(*
SPDX-FileCopyrightText: © 2026 Oleksandr Tiutyk <trofimich@gmail.com>
SPDX-License-Identifier: MIT
License: https://opensource.org/license/mit
*)

(*!
<summary>Base class for one test whose body completes in a single PLC scheduling cycle.</summary>
<description>
Override ExecuteTest with the checks. Returning from the body completes the body automatically.
BeforeTest and AfterTest are optional scenario hooks. Constructor name identifies the case in reports.
Run through TestRunner, directly or inside a TestGroup. A complete run and its reporting may span more cycles
than the body. All instance access belongs to one task without reentry; other tasks need other instances.
</description>
*)

{attribute 'no_explicit_call' := 'do not call this function block directly'}
FUNCTION_BLOCK ABSTRACT SingleCycleTest EXTENDS TestCase

(*!
<summary>Implements the scenario body without runner guards or enumeration.</summary>
<description>
Keep persistent state in instance fields. Reporting a failure does not abort the current callback.
</description>
*)
METHOD PROTECTED ABSTRACT ExecuteTest
END_METHOD

(*!
<summary>Runs the body once and reports completion for the cycle.</summary>
*)
METHOD PROTECTED FINAL RunCycle : TEST_CYCLE_RESULT
ExecuteTest();
RunCycle := TEST_CYCLE_RESULT.DONE;
END_METHOD

END_FUNCTION_BLOCK

(* stored: Version 1.1.0.1
   POU SingleCycleTest: Id {59b4a65d-4a05-4722-819a-36c8562f296a}, SpecialFunc None
   Folder Methods to override: Id {aba7bd54-5472-4bef-8617-736ab163a181}
   Folder Overriden methods: Id {cf9920fa-5d20-449d-822c-735801bafbec}
   Method ExecuteTest: Id {f7894cdc-7848-47ac-aeb9-55a4677731f3}
   Method RunCycle: Id {6045f532-2fae-4f40-9d43-ddf9bb628fbb} *)
